Fanuc KAREL source: KA00137.KL

PROGRAM KA00137
%NOLOCKGROUP
VAR
  SRC: ARRAY[2] OF SHORT
  DST: POSITION
BEGIN
  SRC[1] = 2
  DST = SRC[1]
END KA00137
